Yaskawa INFORM job: RETRACT.JBI

/JOB
//NAME RETRACT
//POS
///NPOS 2,0,0,0,0,0
///TOOL 9
///POSTYPE PULSE
///PULSE
C00000=0,-27,-62,0,46,0
C00001=0,0,0,0,0,0
//INST
///DATE 2026/10/26 01:19
///COMM Generated using RoboDK
///ATTR SC,RW,RJ
///GROUP1 RB1
NOP
'Using Motoman ES200D Base (ta
'rgets wrt base):
'0.0,0.0,0.0,0.0,0.0,0.0
'Setting Tool 9 (USER - CONE -
' 10MM  X  45 DEG):
SETE P00095 (1) 0
SETE P00095 (2) 0
SETE P00095 (3) 85000
SETE P00095 (4) 0
SETE P00095 (5) 0
SETE P00095 (6) 0
SETTOOL TL#(9) P00095
MOVJ C00000 VJ=50.00
MOVJ C00001 VJ=50.00
END
